Universal Robots URScript: Long_ProgramName12.script

def Long_ProgramName12():
  # Default parameters:
  global speed_ms = 0.3
  global speed_rads = 0.75
  global accel_mss = 3
  global accel_radss = 1.2
  global blend_radius_m = 0.001

  # Add subprograms here
  # Start of main program
  # Program generated by RoboDK v5.9.4 for UR10 on 26/10/2026 01:01:20
  # Using nominal kinematics.
  # Long body
  set_tcp(p[0.010000, 0.000000, 0.150000, 0.000000, 0.000000, 0.000000])
  movel([-4.170995, -1.248690, 4.822082, -2.397933, 1.001165, -2.483057],accel_mss,speed_ms,0,blend_radius_m)
  # End of main program
end

Long_ProgramName12()
